PROGRAM Clock
VAR
	{attribute 'hide'} 
	fbClock1OnHz 		: TON;
	{attribute 'hide'} 
	fbClock1OffHz 		: TON;
	{attribute 'hide'} 
	fbClock2OnHz 		: TON;
	{attribute 'hide'} 
	fbClock2OffHz 		: TON;
	{attribute 'hide'} 
	fbClock5OnHz 		: TON;
	{attribute 'hide'} 
	fbClock5OffHz 		: TON;
	{attribute 'hide'} 
	etClockOn2Hz		: TIME;
	{attribute 'hide'} 
	etClockOff2Hz		: TIME;
	{attribute 'hide'} 
	etClockOn1Hz		: TIME;
	{attribute 'hide'} 
	etClockOff1Hz		: TIME;
	{attribute 'hide'} 
	etClockOn5Hz		: TIME;
	{attribute 'hide'} 
	etClockOff5Hz		: TIME;
	pulse1Hz			: BOOL;
	pulse2Hz			: BOOL;
	pulse5Hz			: BOOL;
	{attribute 'hide'} 
	fbClockSr1Hz		: SR;
	{attribute 'hide'} 
	fbClockSr2Hz		: SR;
	{attribute 'hide'} 
	fbClockSr5Hz		: SR;
END_VAR

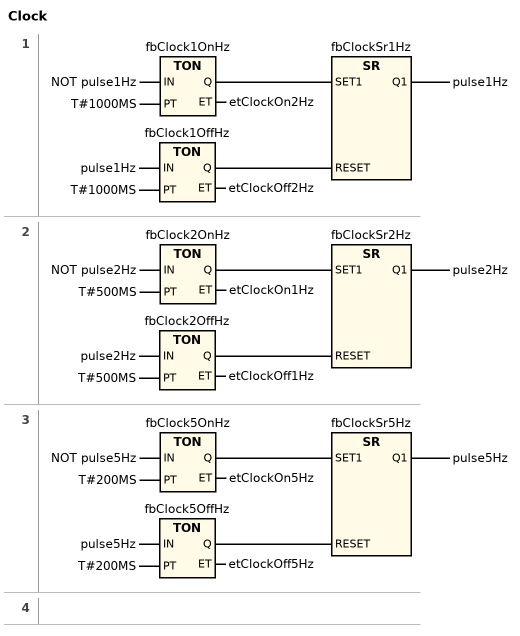
// NETWORK 1
fbClock1OnHz(IN := NOT pulse1Hz, PT := T#1000MS, ET => etClockOn2Hz); // TON
fbClock1OffHz(IN := pulse1Hz, PT := T#1000MS, ET => etClockOff2Hz); // TON
fbClockSr1Hz(SET1 := fbClock1OnHz.Q, RESET := fbClock1OffHz.Q); // SR
pulse1Hz := fbClockSr1Hz.Q1;

// NETWORK 2
fbClock2OnHz(IN := NOT pulse2Hz, PT := T#500MS, ET => etClockOn1Hz); // TON
fbClock2OffHz(IN := pulse2Hz, PT := T#500MS, ET => etClockOff1Hz); // TON
fbClockSr2Hz(SET1 := fbClock2OnHz.Q, RESET := fbClock2OffHz.Q); // SR
pulse2Hz := fbClockSr2Hz.Q1;

// NETWORK 3
fbClock5OnHz(IN := NOT pulse5Hz, PT := T#200MS, ET => etClockOn5Hz); // TON
fbClock5OffHz(IN := pulse5Hz, PT := T#200MS, ET => etClockOff5Hz); // TON
fbClockSr5Hz(SET1 := fbClock5OnHz.Q, RESET := fbClock5OffHz.Q); // SR
pulse5Hz := fbClockSr5Hz.Q1;

// NETWORK 4

END_PROGRAM

(* stored: Version 1.1.0.1, ProductVersion 3.1.4024.12
   POU Clock: Id {541b935e-9f01-46fa-8513-a7a23ad8d0c1}, SpecialFunc None *)
